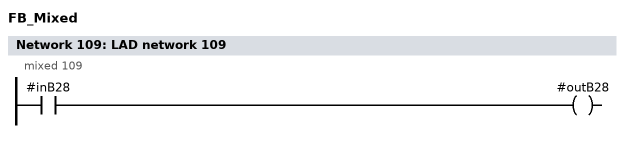
   RUNG wire#powerrail
      Contact( #inB28 )
      Coil( #outB28 )
   END_RUNG
   // the same network as SCL:
   #outB28 := #inB28;
END_REGION

REGION Network 110 (FBD): FBD network 110
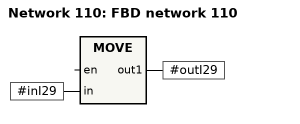
   #outI29 := #inI29;
END_REGION

REGION Network 111 (SCL): SCL network 111
   #tI10 := #inI30 + #cI20;
           IF #inB30 THEN
               #outR10 := #inR10 * 2.0;
           END_IF;
END_REGION

REGION Network 112: LAD network 112
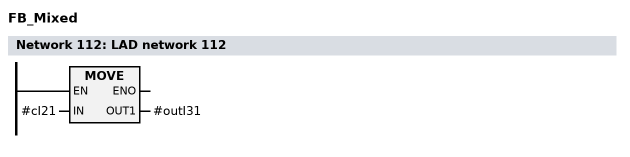
   RUNG wire#powerrail
      Move(in := #cI21, out1 => #outI31)
   END_RUNG
   // the same network as SCL:
   #outI31 := #cI21;
END_REGION

REGION Network 113 (FBD): FBD network 113
   // mixed 113
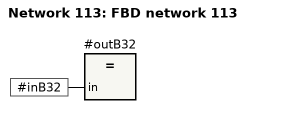
   #outB32 := #inB32;
END_REGION

REGION Network 114 (SCL): SCL network 114
   #tI13 := #inI33 + #cI23;
           IF #inB33 THEN
               #outR13 := #inR13 * 2.0;
           END_IF;
END_REGION

REGION Network 115: LAD network 115
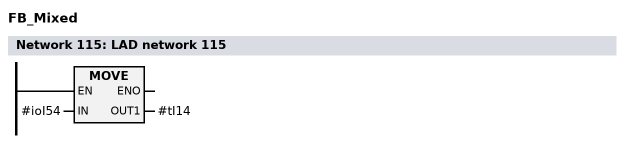
   RUNG wire#powerrail
      Move(in := #ioI54, out1 => #tI14)
   END_RUNG
   // the same network as SCL:
   #tI14 := #ioI54;
END_REGION

REGION Network 116 (FBD): FBD network 116
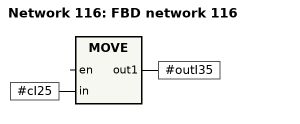
   #outI35 := #cI25;
END_REGION

REGION Network 117 (SCL): SCL network 117
   // mixed 117
   #tI16 := #inI36 + #cI26;
           IF #inB36 THEN
               #outR16 := #inR16 * 2.0;
           END_IF;
END_REGION

REGION Network 118: LAD network 118
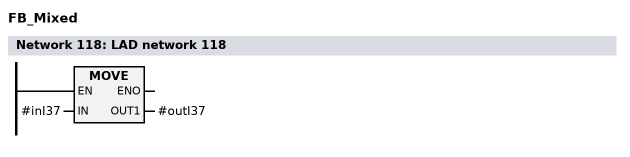
   RUNG wire#powerrail
      Move(in := #inI37, out1 => #outI37)
   END_RUNG
   // the same network as SCL:
   #outI37 := #inI37;
END_REGION

REGION Network 119 (FBD): FBD network 119
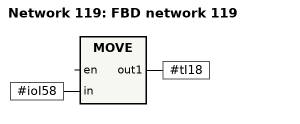
   #tI18 := #ioI58;
END_REGION

REGION Network 120 (SCL): SCL network 120
   #tI19 := #inI39 + #cI29;
           IF #inB39 THEN
               #outR19 := #inR19 * 2.0;
           END_IF;
END_REGION
END_FUNCTION_BLOCK
